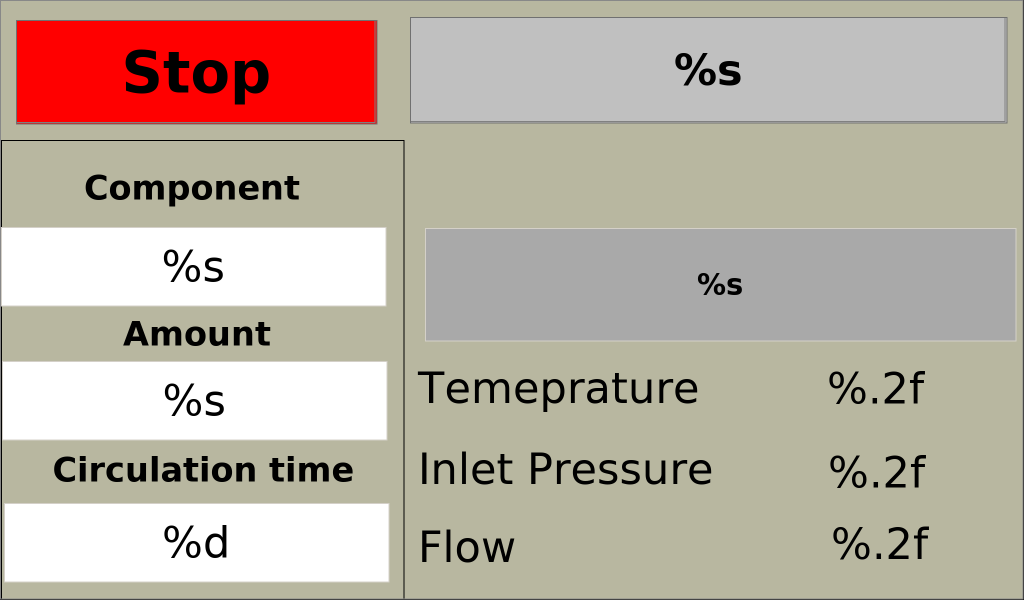
VISUALIZATION Main  // 1024x600
    Rectangle (0,0 1024x600)
    Button (16,20 361x104), "Stop"
    Button (410,17 597x106), "%s", text variable: prg_TriBlender.sStateDescription, input disabled if: prg_TriBlender.bDisableButton
        p2175578022: prg_TriBlender.wButtonColor
        OnMouseClick: execute { prg_TriBlender.bContinue:=TRUE; }
    Rectangle (1,140 403x460)
    Textfield (9,144 378x87), "Component", invisible if: prg_TriBlender.bDisableName
    Textfield (1,227 385x79), "%s", text variable: prg_TriBlender.stTriblender.sComponenetName, invisible if: prg_TriBlender.bDisableName
    Textfield (2,361 385x79), "%s", text variable: prg_TriBlender.stTriblender.sComponenetAmount, invisible if: prg_TriBlender.bDisableAmount
    Textfield (4,302 386x63), "Amount", invisible if: prg_TriBlender.bDisableAmount
    Textfield (7,441 393x57), "Circulation time", invisible if: prg_TriBlender.bDisableTime
    Textfield (4,503 385x79), "%d", text variable: prg_TriBlender.iCirculationTimeLeft, invisible if: prg_TriBlender.bDisableTime
    Textfield (425,228 591x113), "%s", text variable: prg_TriBlender.sStateInstructions
    Textfield (415,444 354x50), "Inlet Pressure"
    Textfield (765,441 223x63), "%.2f", text variable: prg_TriBlender.stTriblender.rPressure
    Textfield (415,522 354x50), "Flow"
    Textfield (767,517 225x54), "%.2f", text variable: prg_TriBlender.stTriblender.rFlow
    Textfield (415,363 354x50), "Temeprature"
    Textfield (764,365 223x47), "%.2f", text variable: prg_TriBlender.stTriblender.rTemp
END_VISUALIZATION

(* stored: Version 1.1.0.1, ProductVersion 3.1.4024.13
   Visu Main: Id {e2a51372-7a75-4142-88f8-0cd1be4fcb07} *)
